(* IEC 61131-3 sources: SemaPLC/sema-plc-benchmark/spec2control-benchmark/data/st-baseline/benzene-distillation/pous/programs, 5 files *)

(* ---- main.st ---- *)
PROGRAM main
VAR
	Heartbeat : bool;
END_VAR

(* Entry point required by OpenPLC Editor v4. The process sections run as parallel program instances under task0; main only provides a scan heartbeat. *)
Heartbeat := NOT Heartbeat;

END_PROGRAM

(* ---- Section2.st ---- *)
PROGRAM Section2
VAR
	TE101_Temperature_PV : real;
	LIT101_Level_PV : real;
	PIT102_Pressure_PV : real;
	TIC104_MV_Percent : real;
	PV103_Position_FB : real;
	TE_101 : ANALOG_IN;
	LIT_101 : ANALOG_IN;
	PIT_102 : ANALOG_IN;
	TIC_104 : PID_BASIC;
	PV_103 : VALVE_ELECTRIC;
	XV_105 : VALVE_ON_OFF;
	LAH_101 : DIGITAL_IN;
	LAL_101 : DIGITAL_IN;
	XV105_NotOpen_NOT : bool;
	TIC104_Inhibit_OR : bool;
	LA_LevelTrip_OR : bool;
END_VAR

TE_101(
    Scaling_Slope := 9.375,
    Scaling_Offset := 12.5,
    Alarm_Enable := TRUE);
LIT_101(
    PV_High := 80.0,
    PV_Low := 20.0,
    Alarm_Enable := TRUE);
PIT_102(
    Alarm_Enable := TRUE);
PV_103(
    Control_Signal := TIC_104.XOUT,
    Open_Limit := 100.0,
    Close_Limit := 0.0);
LAH_101();
LAL_101();
LA_LevelTrip_OR := LAH_101.DI_Out OR LAL_101.DI_Out;
XV_105(
    Inhibit := LA_LevelTrip_OR);
XV105_NotOpen_NOT := NOT XV_105.FB_Opened;
TIC104_Inhibit_OR := PIT_102.High_Alarm OR PIT_102.Low_Alarm OR TE_101.High_Alarm OR TE_101.Low_Alarm OR TE_101.General_Fault OR LIT_101.High_Alarm OR LIT_101.Low_Alarm OR XV105_NotOpen_NOT OR PV_103.Alarm;
TIC_104(
    PV := TE_101.PV,
    SP := 150.0,
    MV_MIN := 10.0,
    MV_MAX := 90.0,
    KP := 3.0,
    TR := 0.5,
    TD := 0.1,
    PV_High := 180.0,
    PV_Low := 130.0,
    Inhibit := TIC104_Inhibit_OR);

(* Outputs published to other sections / HMI. *)
TE101_Temperature_PV := TE_101.PV;
LIT101_Level_PV := LIT_101.PV;
PIT102_Pressure_PV := PIT_102.PV;
TIC104_MV_Percent := TIC_104.XOUT;
PV103_Position_FB := PV_103.Feedback_Pos;

END_PROGRAM

(* ---- Section3.st ---- *)
PROGRAM Section3
VAR
	Reboiler_Temperature_PV_TI106 : real;
	Steam_Flow_PV_FIT101 : real;
	Column_Pressure_PV_PT101 : real;
	FIC104_MV_SteamValveCmd : real;
	LIC002_LowLevel_Trip : bool;
	TI_106 : ANALOG_IN;
	FIT_101 : ANALOG_IN;
	PT_101 : ANALOG_IN;
	FIC_104 : PID_BASIC;
	TCV_106 : VALVE_ELECTRIC;
	LIC_002 : BOOL_INPUT;
	TAH_106 : BOOL_INPUT;
	TAL_106 : BOOL_INPUT;
	FAH_104 : BOOL_INPUT;
	ReboilerTrip_OR : bool;
END_VAR

TI_106(
    PV_High := 190.0,
    PV_Low := 170.0,
    Scaling_Slope := 9.375,
    Scaling_Offset := 62.5,
    Alarm_Enable := TRUE);
FIT_101(
    PV_Low := 10.0,
    Alarm_Enable := TRUE);
PT_101(
    Alarm_Enable := TRUE);
LIC_002(
    Bool_In := LIC002_LowLevel_Trip,
    Alarm_OnTrue := TRUE);
ReboilerTrip_OR := LIC_002.Bool_Out OR FIC_104.PV_High_Alarm OR TI_106.General_Fault OR PT_101.Low_Alarm;
TCV_106(
    Control_Signal := FIC_104.XOUT,
    Manual_Mode := FALSE,
    Manual_Position := 0.0,
    Open_Limit := 100.0,
    Close_Limit := 0.0,
    Inhibit := ReboilerTrip_OR);
FIC_104(
    AUTO := TRUE,
    PV := TI_106.PV,
    SP := 180.0,
    MV_MIN := 0.0,
    MV_MAX := 100.0,
    X0 := TCV_106.Feedback_Pos,
    KP := 3.0,
    TR := 1.2,
    TD := 0.3,
    Inhibit := ReboilerTrip_OR);
TAH_106(
    Bool_In := TI_106.High_Alarm,
    Alarm_OnTrue := TRUE);
TAL_106(
    Bool_In := TI_106.Low_Alarm,
    Alarm_OnTrue := TRUE);
FAH_104(
    Bool_In := FIT_101.Low_Alarm,
    Alarm_OnTrue := TRUE);

(* Outputs published to other sections / HMI. *)
Reboiler_Temperature_PV_TI106 := TI_106.PV;
Steam_Flow_PV_FIT101 := FIT_101.PV;
Column_Pressure_PV_PT101 := PT_101.PV;
FIC104_MV_SteamValveCmd := FIC_104.XOUT;

END_PROGRAM

(* ---- Section4.st ---- *)
PROGRAM Section4
VAR
	LT_105_Level_PV : real;
	FT_107_Flow_PV : real;
	PT_104_Pressure_PV : real;
	LIC_104_RSP_to_FIC_107_GPM : real;
	FIC_107_Control_Signal_to_LV_107 : real;
	XV103_NotOpen : bool;
	Cascade_Inhibit : bool;
	Permissive_OK : bool;
	LT_105 : ANALOG_IN;
	FT_107 : ANALOG_IN;
	PT_104 : ANALOG_IN;
	LIC_104 : PID_BASIC;
	FIC_107 : PID_BASIC;
	PIC_104 : PID_BASIC;
	LV_107 : VALVE_ELECTRIC;
	XV_103 : VALVE_ON_OFF;
	CascadeStartDelay_TON : TON;
	CascadeInhibit_OR : bool;
	XV103NotOpen_NOT : bool;
	CascadePermissive_NOT : bool;
	LIC_to_FIC_SP_MULT : real;
END_VAR

LT_105(
    Alarm_Enable := TRUE);
FT_107(
    Alarm_Enable := TRUE);
PT_104(
    PV_High := 30.0,
    Alarm_Enable := TRUE);
LIC_to_FIC_SP_MULT := LIC_104.XOUT * 0.5;
FIC_107(
    AUTO := Permissive_OK,
    PV := FT_107.PV,
    SP := LIC_to_FIC_SP_MULT,
    MV_MIN := 0.0,
    MV_MAX := 100.0,
    KP := 4.0,
    TR := 0.5,
    TD := 0.0,
    Inhibit := CascadeInhibit_OR);
LV_107(
    Control_Signal := FIC_107.XOUT,
    Manual_Mode := PT_104.High_Alarm,
    Manual_Position := 0.0,
    Open_Limit := 100.0,
    Close_Limit := 0.0,
    Inhibit := PT_104.High_Alarm);
XV_103();
XV103NotOpen_NOT := NOT XV_103.FB_Opened;
CascadeInhibit_OR := XV103NotOpen_NOT OR LT_105.Low_Alarm OR PT_104.Low_Alarm OR PT_104.High_Alarm OR FT_107.General_Fault OR LV_107.Alarm;
CascadeStartDelay_TON(
    IN := Permissive_OK,
    PT := T#30s);
LIC_104(
    AUTO := CascadeStartDelay_TON.Q,
    PV := LT_105.PV,
    SP := 65.0,
    MV_MIN := 0.0,
    MV_MAX := 100.0,
    X0 := 40.0,
    KP := 1.5,
    TR := 2.5,
    TD := 0.0,
    PV_High := 90.0,
    PV_Low := 10.0,
    Inhibit := CascadeInhibit_OR);
PIC_104(
    PV := PT_104.PV);
CascadePermissive_NOT := NOT Cascade_Inhibit;

(* Outputs published to other sections / HMI. *)
LT_105_Level_PV := LT_105.PV;
FT_107_Flow_PV := FT_107.PV;
PT_104_Pressure_PV := PT_104.PV;
LIC_104_RSP_to_FIC_107_GPM := LIC_to_FIC_SP_MULT;
FIC_107_Control_Signal_to_LV_107 := FIC_107.XOUT;
XV103_NotOpen := XV103NotOpen_NOT;
Cascade_Inhibit := CascadeInhibit_OR;
Permissive_OK := CascadePermissive_NOT;

END_PROGRAM

(* ---- Section6.st ---- *)
PROGRAM Section6
VAR
	FT105_FeedFlowRate : real;
	FT106_BottomsFlowRate : real;
	FT106_SP_From_IIC104 : real;
	LIC002_LevelPV : real;
	FT_105 : ANALOG_IN;
	FT_106 : ANALOG_IN;
	FV_101 : VALVE_ELECTRIC;
	IIC_104 : RATIO_CONTROL;
	FIC_106 : PID_BASIC;
	LIC_002 : PID_BASIC;
	LIC_002_LOW_LEVEL_ILK : BOOL_INPUT;
	FEED_PUMP_RUN : DIGITAL_IN;
	BOTTOMS_PUMP_RUN : DIGITAL_IN;
	FeedAboveCutoff_GT : bool;
	PumpsRunning_AND : bool;
	PumpsNotRunning_NOT : bool;
	RatioInhibit_OR : bool;
END_VAR

FT_105(
    PV_Low := 50.0,
    Scaling_Slope := 62.5,
    Scaling_Offset := -250.0,
    Alarm_Enable := TRUE);
FT_106(
    Scaling_Slope := 62.5,
    Scaling_Offset := -250.0,
    Alarm_Enable := TRUE);
FeedAboveCutoff_GT := (FT_105.PV > 50.0);
BOTTOMS_PUMP_RUN();
FEED_PUMP_RUN();
LIC_002(
    PV := LIC002_LevelPV);
LIC_002_LOW_LEVEL_ILK(
    Bool_In := LIC_002.PV_Low_Alarm,
    Alarm_OnTrue := TRUE);
PumpsRunning_AND := FEED_PUMP_RUN.DI_Out AND BOTTOMS_PUMP_RUN.DI_Out;
PumpsNotRunning_NOT := NOT PumpsRunning_AND;
RatioInhibit_OR := LIC_002_LOW_LEVEL_ILK.Bool_Out OR PumpsNotRunning_NOT OR FT_105.General_Fault OR FT_106.General_Fault OR FEED_PUMP_RUN.Fault_State OR BOTTOMS_PUMP_RUN.Fault_State;
IIC_104(
    Auto := FeedAboveCutoff_GT,
    PrimaryPV := FT_105.PV,
    SecondaryPV := FT_106.PV,
    RatioSP := 1.5,
    MV_MIN := 0.0,
    MV_MAX := 1000.0,
    Inhibit := RatioInhibit_OR);
FIC_106(
    AUTO := FeedAboveCutoff_GT,
    PV := FT_106.PV,
    SP := IIC_104.SlaveSP,
    MV_MIN := 0.0,
    MV_MAX := 100.0,
    Inhibit := RatioInhibit_OR);
FV_101(
    Control_Signal := FIC_106.XOUT,
    Inhibit := RatioInhibit_OR);

(* Outputs published to other sections / HMI. *)
FT105_FeedFlowRate := FT_105.PV;
FT106_BottomsFlowRate := FT_106.PV;
FT106_SP_From_IIC104 := IIC_104.SlaveSP;

END_PROGRAM
